(* IEC 61131-3 sources: STruCpp/tests/st-validation/expressions, 8 files *)

(* ---- arithmetic.st ---- *)
PROGRAM ArithmeticTest
  VAR
    add_result : INT;
    sub_result : INT;
    mul_result : INT;
    div_result : INT;
    mod_result : INT;
    neg_result : INT;
    precedence_result : INT;
    paren_result : INT;
    a : INT;
    b : INT;
  END_VAR

  a := 10;
  b := 3;
  add_result := a + b;
  sub_result := a - b;
  mul_result := a * b;
  div_result := a / b;
  mod_result := a MOD b;
  neg_result := -a;
  precedence_result := a + b * 2;
  paren_result := (a + b) * 2;
END_PROGRAM

(* ---- boolean.st ---- *)
PROGRAM BooleanTest
  VAR
    and_result : BOOL;
    or_result : BOOL;
    not_result : BOOL;
    xor_result : BOOL;
    complex_result : BOOL;
    and_ff : BOOL;
    or_tt : BOOL;
  END_VAR

  and_result := TRUE AND TRUE;
  and_ff := FALSE AND TRUE;
  or_result := FALSE OR TRUE;
  or_tt := TRUE OR TRUE;
  not_result := NOT FALSE;
  xor_result := TRUE XOR FALSE;
  complex_result := (TRUE AND FALSE) OR (NOT FALSE);
END_PROGRAM

(* ---- comparison.st ---- *)
PROGRAM ComparisonTest
  VAR
    eq_true : BOOL;
    eq_false : BOOL;
    neq_true : BOOL;
    lt_true : BOOL;
    lt_false : BOOL;
    gt_true : BOOL;
    le_eq : BOOL;
    le_lt : BOOL;
    ge_eq : BOOL;
    ge_gt : BOOL;
  END_VAR

  eq_true := 5 = 5;
  eq_false := 5 = 6;
  neq_true := 5 <> 6;
  lt_true := 3 < 5;
  lt_false := 5 < 3;
  gt_true := 5 > 3;
  le_eq := 5 <= 5;
  le_lt := 3 <= 5;
  ge_eq := 5 >= 5;
  ge_gt := 5 >= 3;
END_PROGRAM

(* ---- test_arithmetic.st ---- *)
TEST 'Addition'
  VAR uut : ArithmeticTest; END_VAR
  uut();
  ASSERT_EQ(uut.add_result, 13);
END_TEST

TEST 'Subtraction'
  VAR uut : ArithmeticTest; END_VAR
  uut();
  ASSERT_EQ(uut.sub_result, 7);
END_TEST

TEST 'Multiplication'
  VAR uut : ArithmeticTest; END_VAR
  uut();
  ASSERT_EQ(uut.mul_result, 30);
END_TEST

TEST 'Integer division truncates'
  VAR uut : ArithmeticTest; END_VAR
  uut();
  ASSERT_EQ(uut.div_result, 3);
END_TEST

TEST 'Modulo operation'
  VAR uut : ArithmeticTest; END_VAR
  uut();
  ASSERT_EQ(uut.mod_result, 1);
END_TEST

TEST 'Unary negation'
  VAR uut : ArithmeticTest; END_VAR
  uut();
  ASSERT_EQ(uut.neg_result, -10);
END_TEST

TEST 'Operator precedence: multiply before add'
  VAR uut : ArithmeticTest; END_VAR
  uut();
  ASSERT_EQ(uut.precedence_result, 16);
END_TEST

TEST 'Parentheses override precedence'
  VAR uut : ArithmeticTest; END_VAR
  uut();
  ASSERT_EQ(uut.paren_result, 26);
END_TEST

(* ---- test_boolean.st ---- *)
TEST 'AND: TRUE AND TRUE = TRUE'
  VAR uut : BooleanTest; END_VAR
  uut();
  ASSERT_TRUE(uut.and_result);
END_TEST

TEST 'AND: FALSE AND TRUE = FALSE'
  VAR uut : BooleanTest; END_VAR
  uut();
  ASSERT_FALSE(uut.and_ff);
END_TEST

TEST 'OR: FALSE OR TRUE = TRUE'
  VAR uut : BooleanTest; END_VAR
  uut();
  ASSERT_TRUE(uut.or_result);
END_TEST

TEST 'OR: TRUE OR TRUE = TRUE'
  VAR uut : BooleanTest; END_VAR
  uut();
  ASSERT_TRUE(uut.or_tt);
END_TEST

TEST 'NOT: NOT FALSE = TRUE'
  VAR uut : BooleanTest; END_VAR
  uut();
  ASSERT_TRUE(uut.not_result);
END_TEST

TEST 'XOR: TRUE XOR FALSE = TRUE'
  VAR uut : BooleanTest; END_VAR
  uut();
  ASSERT_TRUE(uut.xor_result);
END_TEST

TEST 'Complex: (TRUE AND FALSE) OR (NOT FALSE) = TRUE'
  VAR uut : BooleanTest; END_VAR
  uut();
  ASSERT_TRUE(uut.complex_result);
END_TEST

(* ---- test_comparison.st ---- *)
TEST 'Equal: 5 = 5'
  VAR uut : ComparisonTest; END_VAR
  uut();
  ASSERT_TRUE(uut.eq_true);
END_TEST

TEST 'Not equal: 5 = 6 is FALSE'
  VAR uut : ComparisonTest; END_VAR
  uut();
  ASSERT_FALSE(uut.eq_false);
END_TEST

TEST 'Not equal operator: 5 <> 6'
  VAR uut : ComparisonTest; END_VAR
  uut();
  ASSERT_TRUE(uut.neq_true);
END_TEST

TEST 'Less than: 3 < 5'
  VAR uut : ComparisonTest; END_VAR
  uut();
  ASSERT_TRUE(uut.lt_true);
END_TEST

TEST 'Less than false: 5 < 3'
  VAR uut : ComparisonTest; END_VAR
  uut();
  ASSERT_FALSE(uut.lt_false);
END_TEST

TEST 'Greater than: 5 > 3'
  VAR uut : ComparisonTest; END_VAR
  uut();
  ASSERT_TRUE(uut.gt_true);
END_TEST

TEST 'Less or equal when equal: 5 <= 5'
  VAR uut : ComparisonTest; END_VAR
  uut();
  ASSERT_TRUE(uut.le_eq);
END_TEST

TEST 'Less or equal when less: 3 <= 5'
  VAR uut : ComparisonTest; END_VAR
  uut();
  ASSERT_TRUE(uut.le_lt);
END_TEST

TEST 'Greater or equal when equal: 5 >= 5'
  VAR uut : ComparisonTest; END_VAR
  uut();
  ASSERT_TRUE(uut.ge_eq);
END_TEST

TEST 'Greater or equal when greater: 5 >= 3'
  VAR uut : ComparisonTest; END_VAR
  uut();
  ASSERT_TRUE(uut.ge_gt);
END_TEST

(* ---- test_type_conversion.st ---- *)
TEST 'INT to REAL conversion'
  VAR uut : TypeConversionTest; END_VAR
  uut();
  ASSERT_NEAR(uut.int_to_real_result, 42.0, 0.001);
END_TEST

TEST 'REAL to INT rounding'
  VAR uut : TypeConversionTest; END_VAR
  uut();
  (* IEC 61131-3: REAL_TO_INT rounds to nearest integer *)
  ASSERT_EQ(uut.real_to_int_result, 4);
END_TEST

TEST 'INT to DINT widening'
  VAR uut : TypeConversionTest; END_VAR
  uut();
  ASSERT_EQ(uut.int_to_dint_result, 42);
END_TEST

TEST 'BOOL to INT'
  VAR uut : TypeConversionTest; END_VAR
  uut();
  ASSERT_EQ(uut.bool_to_int_result, 1);
END_TEST

(* ---- type_conversion.st ---- *)
PROGRAM TypeConversionTest
  VAR
    int_to_real_result : REAL;
    real_to_int_result : INT;
    int_to_dint_result : DINT;
    bool_to_int_result : INT;
    a : INT;
    b : REAL;
  END_VAR

  a := 42;
  b := 3.7;
  int_to_real_result := INT_TO_REAL(a);
  real_to_int_result := REAL_TO_INT(b);
  int_to_dint_result := INT_TO_DINT(a);
  bool_to_int_result := BOOL_TO_INT(TRUE);
END_PROGRAM
